Fanuc TP program (LS listing): Prog_N.LS

/PROG  Prog_N
/ATTR
OWNER		= MNEDITOR;
COMMENT		= "RoboDK sequence";
PROG_SIZE	= 0;
CREATE		= DATE 31-12-14  TIME 12:00:00;
MODIFIED	= DATE 31-12-14  TIME 12:00:00;
FILE_NAME	= Prog_N;
VERSION		= 0;
LINE_COUNT	= 48;
MEMORY_SIZE	= 0;
PROTECT		= READ_WRITE;
TCD:  STACK_SIZE	= 0,
      TASK_PRIORITY	= 50,
      TIME_SLICE	= 0,
      BUSY_LAMP_OFF	= 0,
      ABORT_REQUEST	= 0,
      PAUSE_REQUEST	= 0;
DEFAULT_GROUP	= 1,*,*,*,*;
CONTROL_CODE	= 00000000 00000000;
/MN
   1:  ! Program generated by VerticalBot Studio for Fanuc LR Mate 200 ;
   2:  ! iD on 25/10/2026 12:00:00 ;
   3:  ! Using nominal kinematics. ;
   4:  PR[9,1]=0.000 ;
   5:  PR[9,2]=0.000 ;
   6:  PR[9,3]=0.000 ;
   7:  PR[9,4]=0.000 ;
   8:  PR[9,5]=0.000 ;
   9:  PR[9,6]=0.000 ;
  10:  UFRAME[9]=PR[9] ;
  11:  UFRAME_NUM=9 ;
  12:  PR[9,1]=10.000 ;
  13:  PR[9,2]=0.000 ;
  14:  PR[9,3]=120.000 ;
  15:  PR[9,4]=0.000 ;
  16:  PR[9,5]=15.000 ;
  17:  PR[9,6]=0.000 ;
  18:  UTOOL[9]=PR[9] ;
  19:  UTOOL_NUM=9 ;
  20:J P[1] 20% CNT10 ;
  21:L P[2] 1000mm/sec CNT10 ;
  22:L P[3] 1000mm/sec CNT0 ;
  23:  PAUSE ;
  24:  WAIT  1.50(sec) ;
  25:  MESSAGE[Say "hi" to the operator] ;
  26:  ! A long comment line that exceeds the usual controller limits ;
  27:  ! for comments by far, really ;
  28:  DO[12]=OFF ;
  29:  OUT_A=ON ;
  30:  $WAITTMOUT=1000 ;
  31:  WAIT DI[4]=OFF TIMEOUT, LBL[1] ;
  32:  MESSAGE[Timed out for LBL 1] ;
  33:  PAUSE ;
  34:  LBL[1] ;
  35:  WAIT IN_B=ON ;
  36:  CALL Program_ ;
  37:  PR[9,1]=250.000 ;
  38:  PR[9,2]=300.000 ;
  39:  PR[9,3]=-10.000 ;
  40:  PR[9,4]=0.000 ;
  41:  PR[9,5]=0.000 ;
  42:  PR[9,6]=90.000 ;
  43:  UFRAME[9]=PR[9] ;
  44:  UFRAME_NUM=9 ;
  45:  UTOOL_NUM=7 ;
  46:  ! UT7:10.0,0.0,120.0,0.0,15.0,0.0 ;
  47:L P[4] 1000mm/sec CNT0 ACC100 ;
  48:J P[5] 15% FINE ACC100 ;
/POS
P[1]{
   GP1:
    UF : 9, UT : 9,
	J1=    -20.000 deg,	J2=    10.000 deg,	J3=    -20.000 deg,
	J4=    30.000 deg,	J5=    -40.000 deg,	J6=    50.000 deg
};
P[2]{
   GP1:
    UF : 9, UT : 9,        CONFIG : 'F U T, 0, 0, 0',
	X =   332.153  mm,	Y =  -359.974  mm,	Z =   826.762  mm,
	W =   -51.647 deg,	P =     9.441 deg,	R =  -168.258 deg
};
P[3]{
   GP1:
    UF : 9, UT : 9,        CONFIG : 'F U T, 0, 0, 0',
	X =   286.258  mm,	Y =  -372.547  mm,	Z =   823.386  mm,
	W =   -52.463 deg,	P =     8.848 deg,	R =  -172.388 deg
};
P[4]{
   GP1:
    UF : 9, UT : 7,        CONFIG : 'F U T, 0, 0, 0',
	X =   332.153  mm,	Y =  -359.974  mm,	Z =   826.762  mm,
	W =   -51.647 deg,	P =     9.441 deg,	R =  -168.258 deg
};
P[5]{
   GP1:
    UF : 9, UT : 7,
	J1=    -20.000 deg,	J2=    10.000 deg,	J3=    -20.000 deg,
	J4=    30.000 deg,	J5=    -40.000 deg,	J6=    50.000 deg
};
/END
